(* IEC 61131-3 sources: STBud-for-TwinCAT/samples/SampleSTFiles, 18 files *)

(* ---- ArrayInStruct.st ---- *)
TYPE ST_SensorArray :
STRUCT
    temperatures:ARRAY[1..16] OF REAL;
    pressures:ARRAY[1..8] OF LREAL;
    names:ARRAY[1..16] OF STRING[32];
    statusFlags:ARRAY[1..16] OF BOOL;
END_STRUCT
END_TYPE

(* ---- ComplexStruct.st ---- *)
TYPE ST_MotorCfg :
STRUCT
    name:STRING[32];
    speed:REAL;
    position:ST_Point;
    state:eMotorState;
    limits:ARRAY[0..3] OF REAL;
    enabled:BOOL;
END_STRUCT
END_TYPE

(* ---- ComprehensiveDatatypes.st ---- *)
TYPE ST_TcPOU :
STRUCT
    name:STRING[255];
    id:GUID;
    dataType:eDataType;
    size:DINT;
    flags:DWORD;
    offset:REAL;
    pData:POINTER TO BYTE;
    pNext:REF_TO ST_TcPOU;
    attributes:ARRAY[1..32] OF STRING[64];
    timestamps:ARRAY[1..32] OF DT;
    comment:WSTRING[512];
END_STRUCT
END_TYPE

(* ---- DeepNestedStruct.st ---- *)
TYPE ST_RobotArm :
STRUCT
    joints:ARRAY[1..6] OF ST_AxisConfig;
    toolOffset:ST_Point;
    speedOverride:REAL;
    accelOverride:REAL;
    mode:eRobotMode;
    errorCodes:ARRAY[1..10] OF DINT;
    isConnected:BOOL;
    lastUpdate:DT;
END_STRUCT
END_TYPE

(* ---- EnumType.st ---- *)
TYPE eMotorState :
(Idle, Accelerating, Running, Decelerating, Error)
END_TYPE

(* ---- EnumWithValues.st ---- *)
TYPE eAlarmPriority :
(LOW, MEDIUM := 5, HIGH := 10, CRITICAL := 20)
END_TYPE

(* ---- MultiDimArray.st ---- *)
TYPE ST_MultiDimArray :
STRUCT
    grid:ARRAY[1..10, 1..10] OF REAL;
    cube:ARRAY[0..2, 0..2, 0..2] OF DINT;
    names:ARRAY[1..5] OF STRING[20];
END_STRUCT
END_TYPE

(* ---- MultiTypeDeclarations.st ---- *)
TYPE eRobotMode :
(Manual, Auto, Jog, Reference, Error := 99)
END_TYPE

TYPE ST_AxisConfig :
STRUCT
    axisName:STRING[16];
    minPos:REAL;
    maxPos:REAL;
    maxVel:REAL;
    maxAcc:REAL;
    encoderResolution:DINT;
    inverted:BOOL;
END_STRUCT
END_TYPE

(* ---- NestedStructType.st ---- *)
TYPE ST_MotorConfig :
STRUCT
    nominalSpeed:REAL;
    maxSpeed:REAL;
    acceleration:REAL;
    deceleration:REAL;
    direction:DINT;
    enabled:BOOL;
    name:STRING[32];
    position:ST_Point;
END_STRUCT
END_TYPE

(* ---- PointerAndRefType.st ---- *)
TYPE ST_MotorData :
STRUCT
    pPosition:POINTER TO LREAL;
    refVelocity:REF_TO REAL;
    name:STRING[64];
    trajectory:ARRAY[0..99] OF REAL;
END_STRUCT
END_TYPE

(* ---- StructType.st ---- *)
TYPE ST_Point :
STRUCT
    x:REAL;
    y:REAL;
    z:REAL;
END_STRUCT
END_TYPE

(* ---- StructWithEnumAndTime.st ---- *)
TYPE ST_AlarmConfig :
STRUCT
    priority:eAlarmPriority;
    message:STRING[128];
    active:BOOL;
    timestamp:TIME;
    count:DINT;
END_STRUCT
END_TYPE

(* ---- Function.st ---- *)
FUNCTION AddValues : INT
VAR_INPUT
    a : INT;
    b : INT;
END_VAR

AddValues := a + b;

END_FUNCTION

(* ---- ChainedAssignmentAndPointers.st ---- *)
FUNCTION_BLOCK FB_Sample
VAR_INPUT
    p1 : POINTER TO ST_Sample;
END_VAR
VAR
    a       : ST_Sample;
    b       : ST_Sample;
    n       : DINT;
    nPrev   : DINT;
    ton1    : TON;
END_VAR
IF p1 <> 0 THEN
    (* chained assignment: write the source value into two targets at once *)
    a.f1 := b.g.f1 := p1^.f1;
    a.f2 := p1^.f2;
    MEMCPY(destAddr := ADR(a.buf), n := SIZEOF(a.buf), srcAddr := ADR(p1^.buf));
    ton1.IN := a.f2 = nPrev;
    ton1(PT := T#500MS);
    a.bActive := NOT ton1.Q;
    nPrev := a.f2;
ELSE
    p1^.f3 := b.f3 := 0;
END_IF
END_FUNCTION_BLOCK

(* ---- FunctionBlock.st ---- *)
FUNCTION_BLOCK FB_Motor
VAR_INPUT
    speed : INT;
    enable : BOOL;
END_VAR
VAR_OUTPUT
    running : BOOL;
END_VAR
VAR
    internalCounter : INT;
END_VAR

IF enable THEN
    running := TRUE;
    internalCounter := internalCounter + speed;
ELSE
    running := FALSE;
    internalCounter := 0;
END_IF;

END_FUNCTION_BLOCK

(* ---- PIDController.st ---- *)
FUNCTION_BLOCK FB_PDController
VAR_INPUT
    setpoint : REAL;
    actualValue : REAL;
    kp : REAL := 1.0;
    ki : REAL := 0.1;
    kd : REAL := 0.01;
    enable : BOOL;
END_VAR
VAR_OUTPUT
    output : REAL;
    error : REAL;
    saturated : BOOL;
END_VAR
VAR
    integral : REAL;
    prevError : REAL;
    dt : TIME := T#10ms;
    maxOutput : REAL := 100.0;
    minOutput : REAL := -100.0;
END_VAR

IF enable THEN
    error := setpoint - actualValue;
    integral := integral + error * TIME_TO_REAL(dt);
    output := kp * error + ki * integral + kd * (error - prevError) / TIME_TO_REAL(dt);
    prevError := error;
    IF output > maxOutput THEN
        output := maxOutput;
        saturated := TRUE;
    ELSIF output < minOutput THEN
        output := minOutput;
        saturated := TRUE;
    ELSE
        saturated := FALSE;
    END_IF
ELSE
    output := 0.0;
    integral := 0.0;
    prevError := 0.0;
    error := 0.0;
    saturated := FALSE;
END_IF

END_FUNCTION_BLOCK

(* ---- Sample1.st ---- *)
PROGRAM MainProgram
    VAR
        counter : INT := 0;
        running : BOOL := FALSE;
        timer : TIME := T#0ms;
        message : STRING[80] := 'Hello';
        values : ARRAY[0..9] OF INT;
        fbMotor : FB_Motor;
    END_VAR

    IF running THEN
        counter := counter + 1;
        IF counter > 10 THEN
            running := FALSE;
            counter := 0;
        ELSIF counter > 5 THEN
            timer := T#500ms;
        ELSE
            timer := T#100ms;
        END_IF
    END_IF
    FOR i := 0 TO 9 DO
        values[i] := i * 2;
    END_FOR
    WHILE counter < 100 DO
        counter := counter + 1;
    END_WHILE
    REPEAT
        counter := counter - 1;
    UNTIL counter <= 0
    END_REPEAT
    CASE counter OF
        0: message := 'Zero';
        1 .. 5: message := 'Low';
        6, 7, 8: message := 'Medium';
    ELSE
        message := 'High';
    END_CASE
    fbMotor.Run(speed := 100);
END_PROGRAM

(* ---- TimeDateLiterals.st ---- *)
PROGRAM TimeLiteralShowcase
VAR
    tonDelay   : TON;
    tofDelay   : TOF;
    xTrigger   : BOOL;
    xDone      : BOOL;
    tCycle     : TIME := T#10MS;
    tLong      : TIME := TIME#1D2H3M4S5MS;
    dStart     : DATE := D#2026-01-15;
    todShift   : TOD := TOD#06:30:00;
    dtStamp    : DT := DT#2026-01-15-06:30:00.500;
    tArray     : ARRAY[1..3] OF TIME := [T#1S, T#2S, T#3S];
END_VAR
tonDelay(IN := xTrigger, PT := T#2S);
tofDelay(IN := tonDelay.Q, PT := T#500MS);
xDone := F_Compare(T#1S, tCycle);
IF tonDelay.ET > T#1.5S THEN
    tCycle := T#0S;
END_IF
CASE tCycle OF
    T#10MS:
        xDone := TRUE;
END_CASE
END_PROGRAM
